// TIA Portal V21 export
// export: Created 2026-11-21T16:00:33.6871453Z, ExportSetting WithDefaults, DisplayName Totally Integrated Automation Portal, DisplayVersion V21, DisplayName STEP 7 Professional, DisplayVersion V21, DisplayName STEP 7 Safety, DisplayVersion V21, DisplayName Tech WebApplication, DisplayVersion V21, DisplayName WinCC Basic/Comfort/Advanced, DisplayVersion V21, DisplayName WinCC Unified, DisplayVersion V21
TagTable "Pump"
  PumpSpeed : Int  (%MW10, HMI_Connection_2, 1 s)
  PumpOn : Bool  (%M0.0, HMI_Connection_2, 100 ms)
  Flow : Real  (%MD20, HMI_Connection_2, 500 ms)
  SpeedSetpoint : Int  ()
